Fanuc KAREL source: KA00083.KL

PROGRAM KA00083
%NOLOCKGROUP
VAR
  SRC: XYZWPREXT
  DST: ARRAY[2] OF BYTE
BEGIN
  SRC.X = 1.0
  DST[1] = SRC
END KA00083
